Fanuc KAREL source: KC00050.KL

PROGRAM KC00050
%NOLOCKGROUP
%ENVIRONMENT REGOPE
VAR
  I: INTEGER
  J: INTEGER
  K: INTEGER
  R: REAL
  B: BOOLEAN
  S: STRING[80]
  T: STRING[80]
  P: PATH
  Q: PATH
  AI: ARRAY[8] OF INTEGER
  AB: ARRAY[244] OF BYTE
  XP: XYZWPR
BEGIN
  SET_TPE_POS_REG(I,XP,J)
END KC00050
